FUNCTION_BLOCK FB_Line_Source EXTENDS FB_SFC_Cycle IMPLEMENTS ITF_FB_SFC_Cycle
VAR_INPUT
	valTankA				:	E_Pis_Name	;
	valTankB				:	E_Pis_Name	;
	valTapWater				:	E_Pis_Name	;
	valTapWater_else		:	E_Pis_Name	;
	valTapWater_Drain		:	E_Pis_Name	;	
	valDrain				:	E_Pis_Name	;
	valCIP					:	E_Pis_Name	;
	valCIP_Sel				:	E_Pis_Name	;
	valBlockWater			:	E_Pis_Name	;	
	valWaterSource			:	E_Pis_Name	;
	valWaterSource_Drain	:	E_Pis_Name	;

END_VAR
VAR_OUTPUT
END_VAR
VAR
	eReq				: E_Line_Source;
	eProcess			: E_Line_Source;
	eStatus				: E_Line_Source;
	
	fbPis				: FB_Piston;
	
	stPis_TankA				: REFERENCE TO ST_Piston;
	stPis_TankB				: REFERENCE TO ST_Piston;
	stPis_TapWater			: REFERENCE TO ST_Piston;
	stPis_TapWater_else		: REFERENCE TO ST_Piston;
	stPis_TapWater_Drain	: REFERENCE TO ST_Piston;
	stPis_Drain				: REFERENCE TO ST_Piston;
	stPis_CIP				: REFERENCE TO ST_Piston;
	stPis_CIP_Sel			: REFERENCE TO ST_Piston;
	stPis_BlockWater		: REFERENCE TO ST_Piston;
	stPis_WaterSource		: REFERENCE TO ST_Piston;
	stPis_WaterSource_Drain	: REFERENCE TO ST_Piston;
	
	stPis_Outlet: ST_Piston;
	tonDrainTime: TON;
	ton_TapWaterNotInUse: TON;
	ton_TapWaterDrain_Timeout: TON;
	rt_Req_Reset: R_TRIG;
END_VAR

act_GetReference();

act_Oper();
//IF NOT Init.x THEN
	act_Status();
//END_IF

m_TapWaterNotInUse();

tonDrainTime(PT:=T#1M, IN:=eStatus=E_Line_Source.eDrain AND eReq=E_Line_Target.eNone);
IF tonDrainTime.Q 
AND eReq=E_Line_Source.eNone
AND eProcess=E_Line_Source.eNone
THEN;
	eReq:=E_Line_Source.eClose;
END_IF

m_Request_Reset(memo:=rt_Req_Reset);//

ACTION _aCIP_active:
bStepDone:=FALSE;
IF TRUE 
AND eStatus=E_Line_Source.eCIP
THEN;
	bStepDone:=TRUE;
END_IF
END_ACTION

ACTION _aCIP_entry:
fbPis.m_SetByRecipe(stPis:=stPis_TankA, 			req:=E_Piston_Recipe_State.Release);		
fbPis.m_SetByRecipe(stPis:=stPis_TankB, 			req:=E_Piston_Recipe_State.Release);
fbPis.m_SetByRecipe(stPis:=stPis_TapWater, 			req:=E_Piston_Recipe_State.Release);
fbPis.m_SetByRecipe(stPis:=stPis_TapWater_Drain, 	req:=E_Piston_Recipe_State.Release);
fbPis.m_SetByRecipe(stPis:=stPis_Drain, 			req:=E_Piston_Recipe_State.Act);
fbPis.m_SetByRecipe(stPis:=stPis_CIP, 				req:=E_Piston_Recipe_State.Act);
fbPis.m_SetByRecipe(stPis:=stPis_CIP_Sel,			req:=E_Piston_Recipe_State.Act);
fbPis.m_SetByRecipe(stPis:=stPis_BlockWater, 		req:=E_Piston_Recipe_State.Act);
fbPis.m_SetByRecipe(stPis:=stPis_WaterSource, 		req:=E_Piston_Recipe_State.Release);
fbPis.m_SetByRecipe(stPis:=stPis_WaterSource_Drain, req:=E_Piston_Recipe_State.Release);
END_ACTION

ACTION _aClose_active:
bStepDone:=FALSE;
IF TRUE 
AND eStatus=E_Line_Source.eClose
THEN;
	bStepDone:=TRUE;
END_IF
END_ACTION

ACTION _aClose_entry:
fbPis.m_SetByRecipe(stPis:=stPis_TankA, 			req:=E_Piston_Recipe_State.Release);		
fbPis.m_SetByRecipe(stPis:=stPis_TankB, 			req:=E_Piston_Recipe_State.Release);
fbPis.m_SetByRecipe(stPis:=stPis_TapWater, 			req:=E_Piston_Recipe_State.Release);
fbPis.m_SetByRecipe(stPis:=stPis_TapWater_Drain, 	req:=E_Piston_Recipe_State.Release);
fbPis.m_SetByRecipe(stPis:=stPis_Drain, 			req:=E_Piston_Recipe_State.Release);
fbPis.m_SetByRecipe(stPis:=stPis_CIP, 				req:=E_Piston_Recipe_State.Release);
fbPis.m_SetByRecipe(stPis:=stPis_CIP_Sel,			req:=E_Piston_Recipe_State.Release);
fbPis.m_SetByRecipe(stPis:=stPis_BlockWater, 		req:=E_Piston_Recipe_State.Release);
fbPis.m_SetByRecipe(stPis:=stPis_WaterSource, 		req:=E_Piston_Recipe_State.Release);
fbPis.m_SetByRecipe(stPis:=stPis_WaterSource_Drain, req:=E_Piston_Recipe_State.Release);
END_ACTION

ACTION _aDone_entry:
eProcess:=E_Line_Source.eNone;
eReq:=E_Line_Source.eNone;
bRun:=FALSE;
bDone:=TRUE;
END_ACTION

ACTION _aDrain_active:
bStepDone:=FALSE;
IF TRUE 
AND eStatus=E_Line_Source.eDrain
THEN;
	bStepDone:=TRUE;
END_IF
END_ACTION

ACTION _aDrain_entry:
fbPis.m_SetByRecipe(stPis:=stPis_TankA, 			req:=E_Piston_Recipe_State.Release);		
fbPis.m_SetByRecipe(stPis:=stPis_TankB, 			req:=E_Piston_Recipe_State.Release);
fbPis.m_SetByRecipe(stPis:=stPis_TapWater, 			req:=E_Piston_Recipe_State.Release);
fbPis.m_SetByRecipe(stPis:=stPis_TapWater_Drain, 	req:=E_Piston_Recipe_State.Release);
fbPis.m_SetByRecipe(stPis:=stPis_Drain, 			req:=E_Piston_Recipe_State.Act);
fbPis.m_SetByRecipe(stPis:=stPis_CIP, 				req:=E_Piston_Recipe_State.Release);
fbPis.m_SetByRecipe(stPis:=stPis_CIP_Sel,			req:=E_Piston_Recipe_State.Release);
fbPis.m_SetByRecipe(stPis:=stPis_BlockWater, 		req:=E_Piston_Recipe_State.Release);
fbPis.m_SetByRecipe(stPis:=stPis_WaterSource, 		req:=E_Piston_Recipe_State.Release);
fbPis.m_SetByRecipe(stPis:=stPis_WaterSource_Drain, req:=E_Piston_Recipe_State.Release);
END_ACTION

ACTION _aFill_Water_waiting_active:
bStepDone:=FALSE;
IF TRUE 
AND ton_TapWaterNotInUse.Q
THEN;
	bStepDone:=TRUE;
END_IF
END_ACTION

ACTION _aFillWater_active:
bStepDone:=FALSE;
IF TRUE 
AND eStatus=E_Line_Source.eFillWater
THEN;
	bStepDone:=TRUE;
END_IF
END_ACTION

ACTION _aFillWater_Drain_active:
;
END_ACTION

ACTION _aFillWater_Drain_entry:
fbPis.m_SetByRecipe(stPis:=stPis_TankA, 			req:=E_Piston_Recipe_State.Release);		
fbPis.m_SetByRecipe(stPis:=stPis_TankB, 			req:=E_Piston_Recipe_State.Release);
fbPis.m_SetByRecipe(stPis:=stPis_TapWater, 			req:=E_Piston_Recipe_State.Release);
fbPis.m_SetByRecipe(stPis:=stPis_TapWater_Drain, 	req:=E_Piston_Recipe_State.Release);
fbPis.m_SetByRecipe(stPis:=stPis_Drain, 			req:=E_Piston_Recipe_State.Release);
fbPis.m_SetByRecipe(stPis:=stPis_CIP, 				req:=E_Piston_Recipe_State.Release);
fbPis.m_SetByRecipe(stPis:=stPis_CIP_Sel,			req:=E_Piston_Recipe_State.Release);
fbPis.m_SetByRecipe(stPis:=stPis_BlockWater, 		req:=E_Piston_Recipe_State.Release);
fbPis.m_SetByRecipe(stPis:=stPis_WaterSource, 		req:=E_Piston_Recipe_State.Release);
fbPis.m_SetByRecipe(stPis:=stPis_WaterSource_Drain, req:=E_Piston_Recipe_State.Act);
END_ACTION

ACTION _aFillWater_entry:
fbPis.m_SetByRecipe(stPis:=stPis_TankA, 			req:=E_Piston_Recipe_State.Release);		
fbPis.m_SetByRecipe(stPis:=stPis_TankB, 			req:=E_Piston_Recipe_State.Release);
fbPis.m_SetByRecipe(stPis:=stPis_TapWater, 			req:=E_Piston_Recipe_State.Release);
fbPis.m_SetByRecipe(stPis:=stPis_TapWater_Drain, 	req:=E_Piston_Recipe_State.Release);
fbPis.m_SetByRecipe(stPis:=stPis_Drain, 			req:=E_Piston_Recipe_State.Release);
fbPis.m_SetByRecipe(stPis:=stPis_CIP, 				req:=E_Piston_Recipe_State.Release);
fbPis.m_SetByRecipe(stPis:=stPis_CIP_Sel,			req:=E_Piston_Recipe_State.Release);
fbPis.m_SetByRecipe(stPis:=stPis_BlockWater, 		req:=E_Piston_Recipe_State.Release);
fbPis.m_SetByRecipe(stPis:=stPis_WaterSource, 		req:=E_Piston_Recipe_State.Act);
fbPis.m_SetByRecipe(stPis:=stPis_WaterSource_Drain, req:=E_Piston_Recipe_State.Release);
END_ACTION

ACTION _aInit_active:
SFCReset:=FALSE;
END_ACTION

ACTION _aInit_exit:
eProcess:=E_Line_Source.eNone;
eReq:=E_Line_Source.eNone;
END_ACTION

ACTION _aReady_active:
CASE eReq OF
	E_Line_Source.eClose:;
			IF TRUE THEN;
				eProcess:=E_Line_Source.eClose;
			END_IF

	E_Line_Source.eTank_A:;
			IF TRUE THEN;
				eProcess:=E_Line_Source.eTank_A;
			END_IF	
			
	E_Line_Source.eTank_B:;
			IF TRUE THEN;
				eProcess:=E_Line_Source.eTank_B;
			END_IF	

	E_Line_Source.eTapWater:;
			IF TRUE THEN;
				eProcess:=E_Line_Source.eTapWater;
			END_IF	
			
	E_Line_Source.eFillWater:;
			IF TRUE THEN;
				eProcess:=E_Line_Source.eFillWater;
			END_IF	
			
	E_Line_Source.eCIP:;
			IF TRUE THEN;
				eProcess:=E_Line_Source.eCIP;
			END_IF	
			
	E_Line_Source.eDrain:;
			IF TRUE THEN;
				eProcess:=E_Line_Source.eDrain;
			END_IF			

END_CASE
END_ACTION

ACTION _aReady_exit:
bRun:=TRUE;
bDone:=FALSE;
END_ACTION

ACTION _aTank_A_active:
bStepDone:=FALSE;
IF TRUE 
AND eStatus=E_Line_Source.eTank_A
THEN;
	bStepDone:=TRUE;
END_IF
END_ACTION

ACTION _aTank_A_entry:
fbPis.m_SetByRecipe(stPis:=stPis_TankA, 			req:=E_Piston_Recipe_State.Act);		
fbPis.m_SetByRecipe(stPis:=stPis_TankB, 			req:=E_Piston_Recipe_State.Release);
fbPis.m_SetByRecipe(stPis:=stPis_TapWater, 			req:=E_Piston_Recipe_State.Release);
fbPis.m_SetByRecipe(stPis:=stPis_TapWater_Drain, 	req:=E_Piston_Recipe_State.Release);
fbPis.m_SetByRecipe(stPis:=stPis_Drain, 			req:=E_Piston_Recipe_State.Release);
fbPis.m_SetByRecipe(stPis:=stPis_CIP, 				req:=E_Piston_Recipe_State.Release);
fbPis.m_SetByRecipe(stPis:=stPis_CIP_Sel,			req:=E_Piston_Recipe_State.Release);
fbPis.m_SetByRecipe(stPis:=stPis_BlockWater, 		req:=E_Piston_Recipe_State.Act);
fbPis.m_SetByRecipe(stPis:=stPis_WaterSource, 		req:=E_Piston_Recipe_State.Release);
fbPis.m_SetByRecipe(stPis:=stPis_WaterSource_Drain, req:=E_Piston_Recipe_State.Release);
END_ACTION

ACTION _aTank_B_active:
bStepDone:=FALSE;
IF TRUE 
AND eStatus=E_Line_Source.eTank_B
THEN;
	bStepDone:=TRUE;
END_IF
END_ACTION

ACTION _aTank_B_entry:
fbPis.m_SetByRecipe(stPis:=stPis_TankA, 			req:=E_Piston_Recipe_State.Release);		
fbPis.m_SetByRecipe(stPis:=stPis_TankB, 			req:=E_Piston_Recipe_State.Act);
fbPis.m_SetByRecipe(stPis:=stPis_TapWater, 			req:=E_Piston_Recipe_State.Release);
fbPis.m_SetByRecipe(stPis:=stPis_TapWater_Drain, 	req:=E_Piston_Recipe_State.Release);
fbPis.m_SetByRecipe(stPis:=stPis_Drain, 			req:=E_Piston_Recipe_State.Release);
fbPis.m_SetByRecipe(stPis:=stPis_CIP, 				req:=E_Piston_Recipe_State.Release);
fbPis.m_SetByRecipe(stPis:=stPis_CIP_Sel,			req:=E_Piston_Recipe_State.Release);
fbPis.m_SetByRecipe(stPis:=stPis_BlockWater, 		req:=E_Piston_Recipe_State.Act);
fbPis.m_SetByRecipe(stPis:=stPis_WaterSource, 		req:=E_Piston_Recipe_State.Release);
fbPis.m_SetByRecipe(stPis:=stPis_WaterSource_Drain, 		req:=E_Piston_Recipe_State.Release);
END_ACTION

ACTION _aTap_Water_waiting_active:
bStepDone:=FALSE;
IF TRUE 
AND ton_TapWaterNotInUse.Q
THEN;
	bStepDone:=TRUE;
END_IF
END_ACTION

ACTION _aTapWater_active:
bStepDone:=FALSE;
IF TRUE 
AND eStatus=E_Line_Source.eTapWater
THEN;
	bStepDone:=TRUE;
END_IF
END_ACTION

ACTION _aTapWater_Drain_active:
//fbPis.m_SetByRecipe(stPis:=stPis_TapWater_Drain, 	req:=E_Piston_Recipe_State.Act);
END_ACTION

ACTION _aTapWater_Drain_entry:
fbPis.m_SetByRecipe(stPis:=stPis_TankA, 			req:=E_Piston_Recipe_State.Release);		
fbPis.m_SetByRecipe(stPis:=stPis_TankB, 			req:=E_Piston_Recipe_State.Release);
fbPis.m_SetByRecipe(stPis:=stPis_TapWater, 			req:=E_Piston_Recipe_State.Release);
fbPis.m_SetByRecipe(stPis:=stPis_TapWater_Drain, 	req:=E_Piston_Recipe_State.Act);
fbPis.m_SetByRecipe(stPis:=stPis_Drain, 			req:=E_Piston_Recipe_State.Release);
fbPis.m_SetByRecipe(stPis:=stPis_CIP, 				req:=E_Piston_Recipe_State.Release);
fbPis.m_SetByRecipe(stPis:=stPis_CIP_Sel,			req:=E_Piston_Recipe_State.Release);
fbPis.m_SetByRecipe(stPis:=stPis_BlockWater, 		req:=E_Piston_Recipe_State.Act);
fbPis.m_SetByRecipe(stPis:=stPis_WaterSource, 		req:=E_Piston_Recipe_State.Release);
fbPis.m_SetByRecipe(stPis:=stPis_WaterSource_Drain, req:=E_Piston_Recipe_State.Release);
END_ACTION

ACTION _aTapWater_entry:
fbPis.m_SetByRecipe(stPis:=stPis_TankA, 			req:=E_Piston_Recipe_State.Release);		
fbPis.m_SetByRecipe(stPis:=stPis_TankB, 			req:=E_Piston_Recipe_State.Release);
fbPis.m_SetByRecipe(stPis:=stPis_TapWater, 			req:=E_Piston_Recipe_State.Act);
fbPis.m_SetByRecipe(stPis:=stPis_TapWater_Drain, 	req:=E_Piston_Recipe_State.Release);
fbPis.m_SetByRecipe(stPis:=stPis_Drain, 			req:=E_Piston_Recipe_State.Release);
fbPis.m_SetByRecipe(stPis:=stPis_CIP, 				req:=E_Piston_Recipe_State.Release);
fbPis.m_SetByRecipe(stPis:=stPis_CIP_Sel,			req:=E_Piston_Recipe_State.Release);
fbPis.m_SetByRecipe(stPis:=stPis_BlockWater, 		req:=E_Piston_Recipe_State.Act);
fbPis.m_SetByRecipe(stPis:=stPis_WaterSource, 		req:=E_Piston_Recipe_State.Release);
fbPis.m_SetByRecipe(stPis:=stPis_WaterSource_Drain, req:=E_Piston_Recipe_State.Release);
END_ACTION

ACTION act_GetReference:
m_Set_SFCFlags_Reference();

stPis_TankA				REF= g_Piston.stPis[valTankA];
stPis_TankB				REF= g_Piston.stPis[valTankB];
stPis_TapWater			REF= g_Piston.stPis[valTapWater];
stPis_TapWater_else		REF= g_Piston.stPis[valTapWater_else];
stPis_TapWater_Drain	REF= g_Piston.stPis[valTapWater_Drain];
stPis_BlockWater		REF= g_Piston.stPis[valBlockWater];
stPis_WaterSource		REF= g_Piston.stPis[valWaterSource];
stPis_WaterSource_Drain	REF= g_Piston.stPis[valWaterSource_Drain];
stPis_Drain				REF= g_Piston.stPis[valDrain];
stPis_CIP				REF= g_Piston.stPis[valCIP];
stPis_CIP_Sel			REF= g_Piston.stPis[valCIP_Sel];
END_ACTION

ACTION act_Oper:
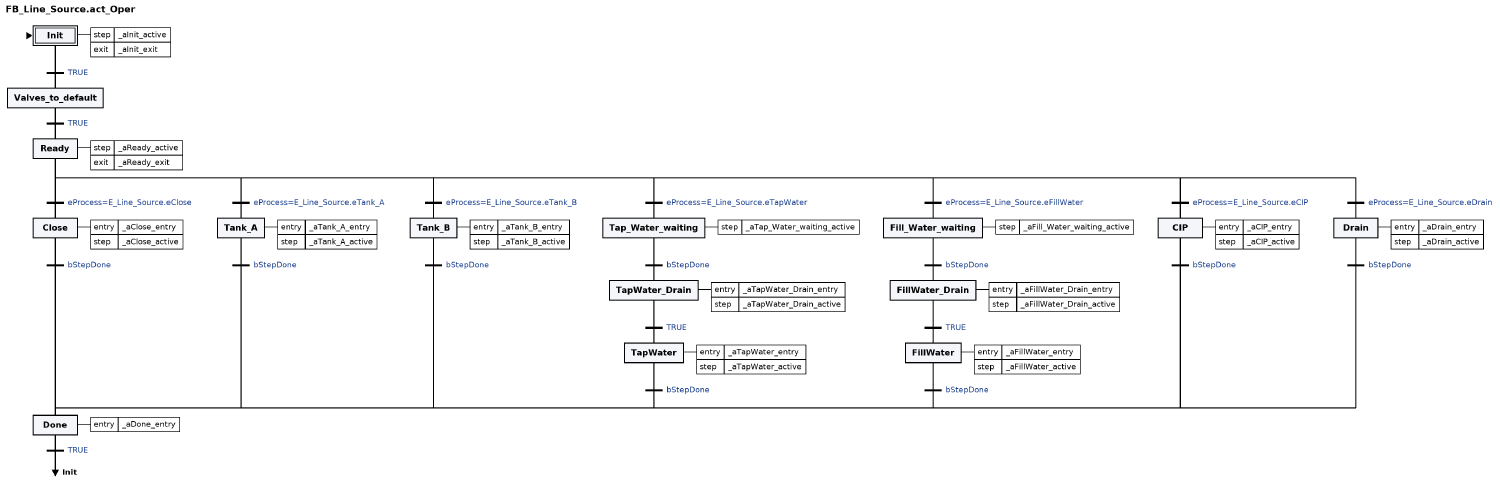
INITIAL_STEP Init:
    _aInit_active(N);  // step action
    _aInit_exit(P0);  // exit action
END_STEP
TRANSITION FROM Init TO Valves_to_default
    := TRUE;
END_TRANSITION
STEP Valves_to_default:
END_STEP
TRANSITION FROM Valves_to_default TO Ready
    := TRUE;
END_TRANSITION
STEP Ready:
    _aReady_active(N);  // step action
    _aReady_exit(P0);  // exit action
END_STEP
TRANSITION FROM Ready TO Close
    := eProcess=E_Line_Source.eClose;
END_TRANSITION
STEP Close:
    _aClose_entry(P1);  // entry action
    _aClose_active(N);  // step action
END_STEP
TRANSITION FROM Close TO Done
    := bStepDone;
END_TRANSITION
TRANSITION FROM Ready TO Tank_A
    := eProcess=E_Line_Source.eTank_A;
END_TRANSITION
STEP Tank_A:
    _aTank_A_entry(P1);  // entry action
    _aTank_A_active(N);  // step action
END_STEP
TRANSITION FROM Tank_A TO Done
    := bStepDone;
END_TRANSITION
TRANSITION FROM Ready TO Tank_B
    := eProcess=E_Line_Source.eTank_B;
END_TRANSITION
STEP Tank_B:
    _aTank_B_entry(P1);  // entry action
    _aTank_B_active(N);  // step action
END_STEP
TRANSITION FROM Tank_B TO Done
    := bStepDone;
END_TRANSITION
TRANSITION FROM Ready TO Tap_Water_waiting
    := eProcess=E_Line_Source.eTapWater;
END_TRANSITION
STEP Tap_Water_waiting:
    _aTap_Water_waiting_active(N);  // step action
END_STEP
TRANSITION FROM Tap_Water_waiting TO TapWater_Drain
    := bStepDone;
END_TRANSITION
STEP TapWater_Drain:  // min time T#10s
    _aTapWater_Drain_entry(P1);  // entry action
    _aTapWater_Drain_active(N);  // step action
END_STEP
TRANSITION FROM TapWater_Drain TO TapWater
    := TRUE;
END_TRANSITION
STEP TapWater:
    _aTapWater_entry(P1);  // entry action
    _aTapWater_active(N);  // step action
END_STEP
TRANSITION FROM TapWater TO Done
    := bStepDone;
END_TRANSITION
TRANSITION FROM Ready TO Fill_Water_waiting
    := eProcess=E_Line_Source.eFillWater;
END_TRANSITION
STEP Fill_Water_waiting:
    _aFill_Water_waiting_active(N);  // step action
END_STEP
TRANSITION FROM Fill_Water_waiting TO FillWater_Drain
    := bStepDone;
END_TRANSITION
STEP FillWater_Drain:  // min time T#10s
    _aFillWater_Drain_entry(P1);  // entry action
    _aFillWater_Drain_active(N);  // step action
END_STEP
TRANSITION FROM FillWater_Drain TO FillWater
    := TRUE;
END_TRANSITION
STEP FillWater:
    _aFillWater_entry(P1);  // entry action
    _aFillWater_active(N);  // step action
END_STEP
TRANSITION FROM FillWater TO Done
    := bStepDone;
END_TRANSITION
TRANSITION FROM Ready TO CIP
    := eProcess=E_Line_Source.eCIP;
END_TRANSITION
STEP CIP:
    _aCIP_entry(P1);  // entry action
    _aCIP_active(N);  // step action
END_STEP
TRANSITION FROM CIP TO Done
    := bStepDone;
END_TRANSITION
TRANSITION FROM Ready TO Drain
    := eProcess=E_Line_Source.eDrain;
END_TRANSITION
STEP Drain:
    _aDrain_entry(P1);  // entry action
    _aDrain_active(N);  // step action
END_STEP
TRANSITION FROM Drain TO Done
    := bStepDone;
END_TRANSITION
STEP Done:
    _aDone_entry(P1);  // entry action
END_STEP
TRANSITION FROM Done TO Init
    := TRUE;
END_TRANSITION
// branch label Branch0_act_Oper
END_ACTION

ACTION act_Status:
IF TRUE 
AND fbPis.m_CheckByRecipe(stPis:=stPis_TankA, 			req:=E_Piston_Recipe_State.Release)		
AND fbPis.m_CheckByRecipe(stPis:=stPis_TankB, 			req:=E_Piston_Recipe_State.Release)
AND fbPis.m_CheckByRecipe(stPis:=stPis_TapWater, 		req:=E_Piston_Recipe_State.Release)
AND fbPis.m_CheckByRecipe(stPis:=stPis_TapWater_Drain, 	req:=E_Piston_Recipe_State.Release)
AND fbPis.m_CheckByRecipe(stPis:=stPis_Drain, 			req:=E_Piston_Recipe_State.Release)
AND fbPis.m_CheckByRecipe(stPis:=stPis_CIP, 			req:=E_Piston_Recipe_State.Release)
AND fbPis.m_CheckByRecipe(stPis:=stPis_CIP_Sel,			req:=E_Piston_Recipe_State.Release)
AND fbPis.m_CheckByRecipe(stPis:=stPis_BlockWater, 		req:=E_Piston_Recipe_State.Release)
AND fbPis.m_CheckByRecipe(stPis:=stPis_WaterSource, 	req:=E_Piston_Recipe_State.Release)
AND fbPis.m_CheckByRecipe(stPis:=stPis_WaterSource_Drain,req:=E_Piston_Recipe_State.Release)
THEN;
	eStatus:=E_Line_Source.eClose;
ELSIF TRUE 
AND fbPis.m_CheckByRecipe(stPis:=stPis_TankA, 			req:=E_Piston_Recipe_State.Act)		
AND fbPis.m_CheckByRecipe(stPis:=stPis_TankB, 			req:=E_Piston_Recipe_State.Release)
AND fbPis.m_CheckByRecipe(stPis:=stPis_TapWater, 		req:=E_Piston_Recipe_State.Release)
AND fbPis.m_CheckByRecipe(stPis:=stPis_TapWater_Drain, 	req:=E_Piston_Recipe_State.Release)
AND fbPis.m_CheckByRecipe(stPis:=stPis_Drain, 			req:=E_Piston_Recipe_State.Release)
AND fbPis.m_CheckByRecipe(stPis:=stPis_CIP, 			req:=E_Piston_Recipe_State.Release)
AND fbPis.m_CheckByRecipe(stPis:=stPis_CIP_Sel,			req:=E_Piston_Recipe_State.Release)
AND fbPis.m_CheckByRecipe(stPis:=stPis_BlockWater, 		req:=E_Piston_Recipe_State.Act)
AND fbPis.m_CheckByRecipe(stPis:=stPis_WaterSource, 	req:=E_Piston_Recipe_State.Release)
AND fbPis.m_CheckByRecipe(stPis:=stPis_WaterSource_Drain,req:=E_Piston_Recipe_State.Release)
THEN;
	eStatus:=E_Line_Source.eTank_A;
ELSIF TRUE 
AND fbPis.m_CheckByRecipe(stPis:=stPis_TankA, 			req:=E_Piston_Recipe_State.Release)		
AND fbPis.m_CheckByRecipe(stPis:=stPis_TankB, 			req:=E_Piston_Recipe_State.Act)
AND fbPis.m_CheckByRecipe(stPis:=stPis_TapWater, 		req:=E_Piston_Recipe_State.Release)
AND fbPis.m_CheckByRecipe(stPis:=stPis_TapWater_Drain, 	req:=E_Piston_Recipe_State.Release)
AND fbPis.m_CheckByRecipe(stPis:=stPis_Drain, 			req:=E_Piston_Recipe_State.Release)
AND fbPis.m_CheckByRecipe(stPis:=stPis_CIP, 			req:=E_Piston_Recipe_State.Release)
AND fbPis.m_CheckByRecipe(stPis:=stPis_CIP_Sel,			req:=E_Piston_Recipe_State.Release)
AND fbPis.m_CheckByRecipe(stPis:=stPis_BlockWater, 		req:=E_Piston_Recipe_State.Act)
AND fbPis.m_CheckByRecipe(stPis:=stPis_WaterSource, 	req:=E_Piston_Recipe_State.Release)
AND fbPis.m_CheckByRecipe(stPis:=stPis_WaterSource_Drain,req:=E_Piston_Recipe_State.Release)
THEN;
	eStatus:=E_Line_Source.eTank_B;
ELSIF TRUE 
AND fbPis.m_CheckByRecipe(stPis:=stPis_TankA, 			req:=E_Piston_Recipe_State.Release)		
AND fbPis.m_CheckByRecipe(stPis:=stPis_TankB, 			req:=E_Piston_Recipe_State.Release)
AND fbPis.m_CheckByRecipe(stPis:=stPis_TapWater, 		req:=E_Piston_Recipe_State.Act)
AND fbPis.m_CheckByRecipe(stPis:=stPis_TapWater_Drain, 	req:=E_Piston_Recipe_State.Release)
AND fbPis.m_CheckByRecipe(stPis:=stPis_TapWater_else, 	req:=E_Piston_Recipe_State.Release)
AND fbPis.m_CheckByRecipe(stPis:=stPis_Drain, 			req:=E_Piston_Recipe_State.Release)
AND fbPis.m_CheckByRecipe(stPis:=stPis_CIP, 			req:=E_Piston_Recipe_State.Release)
AND fbPis.m_CheckByRecipe(stPis:=stPis_CIP_Sel,			req:=E_Piston_Recipe_State.Release)
AND fbPis.m_CheckByRecipe(stPis:=stPis_BlockWater, 		req:=E_Piston_Recipe_State.Act)
AND fbPis.m_CheckByRecipe(stPis:=stPis_WaterSource, 	req:=E_Piston_Recipe_State.Release)
AND fbPis.m_CheckByRecipe(stPis:=stPis_WaterSource_Drain,req:=E_Piston_Recipe_State.Release)
THEN;
	eStatus:=E_Line_Source.eTapWater;
ELSIF TRUE 
AND fbPis.m_CheckByRecipe(stPis:=stPis_TankA, 			req:=E_Piston_Recipe_State.Release)		
AND fbPis.m_CheckByRecipe(stPis:=stPis_TankB, 			req:=E_Piston_Recipe_State.Release)
AND fbPis.m_CheckByRecipe(stPis:=stPis_TapWater, 		req:=E_Piston_Recipe_State.Release)
AND fbPis.m_CheckByRecipe(stPis:=stPis_TapWater_Drain, 	req:=E_Piston_Recipe_State.Release)
AND fbPis.m_CheckByRecipe(stPis:=stPis_Drain, 			req:=E_Piston_Recipe_State.Release)
AND fbPis.m_CheckByRecipe(stPis:=stPis_CIP, 			req:=E_Piston_Recipe_State.Release)
AND fbPis.m_CheckByRecipe(stPis:=stPis_CIP_Sel,			req:=E_Piston_Recipe_State.Release)
AND fbPis.m_CheckByRecipe(stPis:=stPis_BlockWater, 		req:=E_Piston_Recipe_State.Release)
AND fbPis.m_CheckByRecipe(stPis:=stPis_WaterSource, 	req:=E_Piston_Recipe_State.Act)
AND fbPis.m_CheckByRecipe(stPis:=stPis_WaterSource_Drain,req:=E_Piston_Recipe_State.Release)
THEN;
	eStatus:=E_Line_Source.eFillWater;
ELSIF TRUE 
AND fbPis.m_CheckByRecipe(stPis:=stPis_TankA, 			req:=E_Piston_Recipe_State.Release)		
AND fbPis.m_CheckByRecipe(stPis:=stPis_TankB, 			req:=E_Piston_Recipe_State.Release)
AND fbPis.m_CheckByRecipe(stPis:=stPis_TapWater, 		req:=E_Piston_Recipe_State.Release)
AND fbPis.m_CheckByRecipe(stPis:=stPis_TapWater_Drain, 	req:=E_Piston_Recipe_State.Release)
AND fbPis.m_CheckByRecipe(stPis:=stPis_Drain, 			req:=E_Piston_Recipe_State.Act)
AND fbPis.m_CheckByRecipe(stPis:=stPis_CIP, 			req:=E_Piston_Recipe_State.Act)
AND fbPis.m_CheckByRecipe(stPis:=stPis_CIP_Sel,			req:=E_Piston_Recipe_State.Act)
AND fbPis.m_CheckByRecipe(stPis:=stPis_BlockWater, 		req:=E_Piston_Recipe_State.Act)
AND fbPis.m_CheckByRecipe(stPis:=stPis_WaterSource, 	req:=E_Piston_Recipe_State.Release)
AND fbPis.m_CheckByRecipe(stPis:=stPis_WaterSource_Drain,req:=E_Piston_Recipe_State.Release)
THEN;
	eStatus:=E_Line_Source.eCIP;
ELSIF TRUE 
AND fbPis.m_CheckByRecipe(stPis:=stPis_TankA, 			req:=E_Piston_Recipe_State.Release)		
AND fbPis.m_CheckByRecipe(stPis:=stPis_TankB, 			req:=E_Piston_Recipe_State.Release)
AND fbPis.m_CheckByRecipe(stPis:=stPis_TapWater, 		req:=E_Piston_Recipe_State.Release)
AND fbPis.m_CheckByRecipe(stPis:=stPis_TapWater_Drain, 	req:=E_Piston_Recipe_State.Release)
AND fbPis.m_CheckByRecipe(stPis:=stPis_Drain, 			req:=E_Piston_Recipe_State.Act)
AND fbPis.m_CheckByRecipe(stPis:=stPis_CIP, 			req:=E_Piston_Recipe_State.Release)
AND fbPis.m_CheckByRecipe(stPis:=stPis_CIP_Sel,			req:=E_Piston_Recipe_State.Release)
AND fbPis.m_CheckByRecipe(stPis:=stPis_BlockWater, 		req:=E_Piston_Recipe_State.Release)
AND fbPis.m_CheckByRecipe(stPis:=stPis_WaterSource, 	req:=E_Piston_Recipe_State.Release)
AND fbPis.m_CheckByRecipe(stPis:=stPis_WaterSource_Drain,req:=E_Piston_Recipe_State.Release)
THEN;
	eStatus:=E_Line_Source.eDrain;
ELSE;
	eStatus:=E_Line_Source.eNone;
END_IF
END_ACTION

METHOD m_CheckStatus : BOOL
VAR_INPUT
	eReqStatus		: E_Line_Source;
END_VAR
IF eStatus=eReqStatus 
AND eProcess=E_Line_Source.eNone
AND eReq=E_Line_Source.eNone
AND bReady
AND bDone
AND NOT bRun
THEN;
	m_CheckStatus:=TRUE;
END_IF
END_METHOD

METHOD m_Request_Reset : BOOL
VAR_IN_OUT
	memo: R_TRIG;
END_VAR
memo(CLK:=eReq=0);
IF TRUE 
AND memo.Q
THEN;
	SFCReset:=TRUE;
END_IF
END_METHOD

METHOD m_Run : BOOL
VAR_INPUT
	eReqProc			: E_Line_Source;
END_VAR
IF eProcess=E_Line_Source.eNone THEN;
	eProcess:=eReq:=eReqProc;
	bDone:=FALSE;
	m_Run:=TRUE;
END_IF
END_METHOD

METHOD m_Set_SFCFlags_Reference : BOOL
//Set reference to SFC flags

refSFC.SFCInit REF= SFCInit;
refSFC.SFCReset REF= SFCReset;
refSFC.SFCError REF= SFCError;
refSFC.SFCEnableLimit REF= SFCEnableLimit;
refSFC.SFCErrorStep REF= SFCErrorStep;
refSFC.SFCErrorPOU REF= SFCErrorPOU;
refSFC.SFCQuitError REF= SFCQuitError;
refSFC.SFCPause REF= SFCPause;
refSFC.SFCTrans REF= SFCTrans;
refSFC.SFCCurrentStep REF= SFCCurrentStep;
refSFC.SFCTip REF= SFCTip;
refSFC.SFCTipMode REF= SFCTipMode;

// Cycle handle for SFC
m_SFC_Handle();
END_METHOD

METHOD m_TapWaterNotInUse : BOOL
VAR_INPUT
END_VAR
IF TRUE 
AND fbPis.m_CheckByRecipe(stPis:=stPis_TapWater, 			req:=E_Piston_Recipe_State.Release)		
AND fbPis.m_CheckByRecipe(stPis:=stPis_TapWater_Drain, 		req:=E_Piston_Recipe_State.Release)
AND fbPis.m_CheckByRecipe(stPis:=stPis_TapWater_else, 		req:=E_Piston_Recipe_State.Release)
AND fbPis.m_CheckByRecipe(stPis:=stPis_WaterSource, 		req:=E_Piston_Recipe_State.Release)
AND fbPis.m_CheckByRecipe(stPis:=stPis_WaterSource_Drain, 	req:=E_Piston_Recipe_State.Release)
THEN;
	ton_TapWaterNotInUse(IN:=TRUE);
ELSE;
	ton_TapWaterNotInUse(IN:=FALSE);
END_IF

ton_TapWaterNotInUse(PT:=T#3S);


//Tap Water Drain Timeout
ton_TapWaterDrain_Timeout(PT:=T#10S);
IF fbPis.m_CheckByRecipe(stPis:=stPis_TapWater_Drain, 	req:=E_Piston_Recipe_State.Act) THEN;
	ton_TapWaterDrain_Timeout.IN:=TRUE;
ELSE;
	ton_TapWaterDrain_Timeout.IN:=FALSE;
END_IF
IF ton_TapWaterDrain_Timeout.Q THEN;
	fbPis.m_SetByRecipe(stPis:=stPis_TapWater_Drain, 	req:=E_Piston_Recipe_State.Release);
END_IF
END_METHOD

END_FUNCTION_BLOCK

(* stored: Version 1.1.0.1, ProductVersion 3.1.4024.15
   POU FB_Line_Source: Id {137ed242-9f5e-44a3-a945-e1d43cf34d59}, SpecialFunc None
   Folder Manage: Id {88761bd7-027b-418f-9edc-eb285488f960}
   Action _aCIP_active: Id {d20e9967-4c28-47ef-96b1-f277270a5409}
   Action _aCIP_entry: Id {13dab27e-deae-40cd-ac78-cdf4842002bf}
   Action _aClose_active: Id {800028b8-d3dd-442c-9182-b7a96d7ee8e2}
   Action _aClose_entry: Id {182c9ae5-08be-41d6-9707-9097c7820fc5}
   Action _aDone_entry: Id {d5d1f6a7-eea7-4f0a-812c-bd08184c1fb8}
   Action _aDrain_active: Id {b081ccb6-d409-4997-ac13-95a702fa85ab}
   Action _aDrain_entry: Id {abae8c70-1d8c-4cf1-a310-7c62690ed16a}
   Action _aFill_Water_waiting_active: Id {54b5198a-182e-4a0b-a97e-2d5a4448b7f5}
   Action _aFillWater_active: Id {70fede1d-ced9-4535-baf7-250cc6847327}
   Action _aFillWater_Drain_active: Id {c7f0fa82-2cab-4023-89d4-9e59cb147289}
   Action _aFillWater_Drain_entry: Id {a3a1ed40-aff2-4529-a8db-1a966547f62b}
   Action _aFillWater_entry: Id {b4f4e998-dc9c-44aa-b10d-0a06724c51f5}
   Action _aInit_active: Id {391dbbf9-7a55-47eb-943a-cf2da131baa4}
   Action _aInit_exit: Id {935e0fe4-d5a9-42d9-9272-0dadea5e6819}
   Action _aReady_active: Id {0e401379-cf24-47d0-855d-d82202d84006}
   Action _aReady_exit: Id {3c53b576-ca96-486b-88ba-a05f52ed43d6}
   Action _aTank_A_active: Id {cf1041fe-0360-41bb-ac66-2373efb92215}
   Action _aTank_A_entry: Id {ac8bc15e-bac4-4064-93e1-7223870c6aa3}
   Action _aTank_B_active: Id {ad3abc4f-db10-4dca-891a-d858a0ec994e}
   Action _aTank_B_entry: Id {65c0f2c4-cc0b-4481-bd5a-a8dca76e3581}
   Action _aTap_Water_waiting_active: Id {9522d026-ad10-49a7-9cfe-83cab6bca8d4}
   Action _aTapWater_active: Id {0e812b07-28fe-4615-b3fd-f06ab7639658}
   Action _aTapWater_Drain_active: Id {5428fc42-e7f4-4161-852c-f744b46b39f5}
   Action _aTapWater_Drain_entry: Id {d7482c71-9386-488f-9fed-3d026818383a}
   Action _aTapWater_entry: Id {0e5ac7bd-d376-4702-bd92-e1298dc3d345}
   Action act_GetReference: Id {4f2d3bb4-7e54-445d-9be1-c7af3ee92176}
   Action act_Oper: Id {55b69863-d4f1-48da-9cf6-1551e676410b}
   Action act_Status: Id {3024ea02-87ce-4d11-b8f4-5b8eb6467f35}
   Method m_CheckStatus: Id {4048b8d2-9673-4029-84b4-7685ad242031}
   Method m_Request_Reset: Id {a20f9c0a-99d9-433b-80f9-02dafa9d62e9}
   Method m_Run: Id {b3f2817c-37d1-47ea-82d9-76c7c92e82ed}
   Method m_Set_SFCFlags_Reference: Id {1d953b94-b8b7-4eef-b8a4-b7c9f4438caf}
   Method m_TapWaterNotInUse: Id {19fb02a0-95ee-46b4-bcf1-7101cd230b89} *)
